(* IEC 61131-3 sources: beckhoffAutomationInterface/ST/sample, 9 files *)

(* ---- E_MotorState.st ---- *)
{attribute 'qualified_only'}
TYPE E_MotorState :
(
	Idle 		:= 0,
	Running 	:= 1,
	Faulted 	:= 2
);
END_TYPE

(* ---- ST_MotorStatus.st ---- *)
{attribute 'pack_mode' := '1'}
TYPE ST_MotorStatus :
STRUCT
	bRunning 	: BOOL;		// TRUE while the motor is running
	nErrorCode 	: UDINT;	// Non-zero when the motor has faulted
END_STRUCT
END_TYPE

(* ---- T_MotorSpeed.st ---- *)
TYPE T_MotorSpeed : LREAL;
END_TYPE

(* ---- GVL_Shark.st ---- *)
{attribute 'qualified_only'}
VAR_GLOBAL
	nMaxMotorSpeed 	: LREAL 	:= 100.0;	// Global speed limit shared across the project
	sPlantName 		: STRING 	:= 'Shark';	// Human-readable plant/project name
	bMotorRunSensor 	AT %I* 	: BOOL;		// Physical input: motor-running feedback sensor (to be linked to hardware)
	bMotorEnableOutput 	AT %Q* 	: BOOL;		// Physical output: motor enable command (to be linked to hardware)
END_VAR

(* ---- I_Motor.st ---- *)
INTERFACE I_Motor

METHOD Init : BOOL
VAR_INPUT
END_VAR

METHOD Reset : BOOL
VAR_INPUT
END_VAR

(* ---- F_ClampSpeed.st ---- *)
FUNCTION F_ClampSpeed : LREAL
VAR_INPUT
	fSpeed 	: LREAL;	// Requested speed
	fMax 	: LREAL;	// Maximum allowed speed
END_VAR

IF fSpeed > fMax THEN
	F_ClampSpeed := fMax;
ELSE
	F_ClampSpeed := fSpeed;
END_IF

(* ---- FB_Motor.st ---- *)
FUNCTION_BLOCK FB_Motor EXTENDS FB_MotorBase IMPLEMENTS I_Motor
VAR_INPUT
	bStart 	: BOOL;				// Start command
END_VAR
VAR_OUTPUT
	eState 		: E_MotorState;		// Current motor state
	stStatus 	: ST_MotorStatus;	// Current motor status
END_VAR
VAR
	fSpeed 	: T_MotorSpeed := 0;	// Current speed, ramped up while running
END_VAR

// Main cyclic logic of the motor function block
IF bStart THEN
	eState 	:= E_MotorState.Running;
	fSpeed 	:= CalculateRampedSpeed();
ELSE
	eState 	:= E_MotorState.Idle;
	fSpeed 	:= 0;
END_IF

// Drive the physical enable output from the start command, and only report
// "Running" once the physical run-sensor input confirms it
GVL_Shark.bMotorEnableOutput 	:= bStart;
stStatus.bRunning 				:= (eState = E_MotorState.Running) AND GVL_Shark.bMotorRunSensor;
stStatus.nErrorCode := 0;

METHOD PUBLIC Init : BOOL
VAR_INPUT
END_VAR

// One-time initialization, called once from MAIN on the first cycle
fSpeed 	:= 0;
eState 	:= E_MotorState.Idle;
Init 	:= TRUE;

METHOD PUBLIC Reset : BOOL
VAR_INPUT
END_VAR

// Clears speed, state, and status back to defaults
fSpeed 				:= 0;
eState 				:= E_MotorState.Idle;
stStatus.bRunning 	:= FALSE;
stStatus.nErrorCode := 0;
Reset 				:= TRUE;

METHOD PUBLIC Stop : BOOL
VAR_INPUT
END_VAR

// Overrides the abstract FB_MotorBase.Stop \u2014 forces the motor back to idle
eState 				:= E_MotorState.Idle;
fSpeed 				:= 0;
stStatus.bRunning 	:= FALSE;
Stop 				:= TRUE;

METHOD PRIVATE CalculateRampedSpeed : T_MotorSpeed
VAR_INPUT
END_VAR

// Internal helper (not part of I_Motor): ramps fSpeed up by 1.0 each cycle, clamped to 100.0
CalculateRampedSpeed := F_ClampSpeed(fSpeed := fSpeed + 1.0, fMax := 100.0);

(* ---- FB_MotorBase.st ---- *)
{abstract}
FUNCTION_BLOCK FB_MotorBase
VAR
END_VAR

{abstract}
METHOD Stop : BOOL
VAR_INPUT
END_VAR

(* ---- MAIN.st ---- *)
PROGRAM MAIN
VAR
	sHelloWorld 	: STRING 	:= 'Hello, World!'; 	// Sample greeting string
	nCounter		: DINT 		:= 0; 					// Increments once every PLC cycle
	fbMotor			: FB_Motor;							// Motor function block instance
	ipMotor			: I_Motor;							// Interface reference to fbMotor, exercised via I_Motor
	bInitDone		: BOOL 		:= FALSE;				// Latches once Init() has run
	bResetDone		: BOOL 		:= FALSE;				// Latches the result of the last Reset() call
	bStopDone		: BOOL 		:= FALSE;				// Latches the result of the last Stop() call
END_VAR

// Increment the counter on every cycle
nCounter := nCounter + 1;

// Bind the interface reference to the FB instance (FB_Motor IMPLEMENTS I_Motor)
ipMotor := fbMotor;

// Call Init() once on the first cycle, via the interface
IF NOT bInitDone THEN
	bInitDone := ipMotor.Init();
END_IF

// Periodically reset the motor (demo trigger), via the interface
IF nCounter MOD 1000 = 0 THEN
	bResetDone := ipMotor.Reset();
END_IF

// Periodically stop the motor (demo trigger), calling the overridden
// FB_MotorBase.Stop directly on the instance (Stop is not part of I_Motor)
IF nCounter MOD 5000 = 0 THEN
	bStopDone := fbMotor.Stop();
END_IF

// Drive the motor and run its main cyclic logic
fbMotor(bStart := TRUE);
